// TIA Portal V20 export
Screen "Pop-up_Hmi_Opmodes18_h_Popup"  585x540
  ScreenItem "Background" at 0,0 size 585x540  Type=HmiRectangle
  ScreenItem "Dummy8" at 293,111 size 25x25  Type=HmiRectangle
  ScreenItem "Dummy9" at 319,111 size 25x25  Type=HmiRectangle
  ScreenItem "Dummy10" at 345,111 size 25x25  Type=HmiRectangle
  ScreenItem "Dummy11" at 371,111 size 25x25  Type=HmiRectangle
  ScreenItem "Dummy12" at 397,111 size 25x25  Type=HmiRectangle
  ScreenItem "Textfeld_1" at 77,106 size 29x30  Type=HmiTextBox
  ScreenItem "Dummy6" at 241,111 size 25x25  Type=HmiRectangle
  ScreenItem "Text_HmiPanelNo" at 244,50 size 160x23  Type=HmiTextBox
  ScreenItem "State_OPMode8_Select" at 293,80 size 25x25  Type=HmiTextBox
  ScreenItem "State_OPMode8_NotSelect" at 293,80 size 25x25  Type=HmiTextBox
  ScreenItem "State_OPMode8_Vis" at 293,80 size 25x25  Type=HmiRectangle
  ScreenItem "Descr_OPMode" at 108,26 size 305x20  Type=HmiTextBox
  ScreenItem "Dummy7" at 267,111 size 25x25  Type=HmiRectangle
  ScreenItem "Overview_OPMode" at 1,1 size 519x25  Type=HmiTextBox
  ScreenItem "State_OPMode1_Select" at 111,80 size 25x25  Type=HmiTextBox
  ScreenItem "State_OPMode1_NotSelect" at 111,80 size 25x25  Type=HmiTextBox
  ScreenItem "State_OPMode1_Vis" at 111,80 size 25x25  Type=HmiRectangle
  ScreenItem "State_OPMode2_Select" at 137,80 size 25x25  Type=HmiTextBox
  ScreenItem "State_OPMode2_NotSelect" at 137,80 size 25x25  Type=HmiTextBox
  ScreenItem "State_OPMode2_Vis" at 137,80 size 25x25  Type=HmiRectangle
  ScreenItem "State_OPMode3_Select" at 163,80 size 25x25  Type=HmiTextBox
  ScreenItem "State_OPMode3_NotSelect" at 163,80 size 25x25  Type=HmiTextBox
  ScreenItem "State_OPMode3_Vis" at 163,80 size 25x25  Type=HmiRectangle
  ScreenItem "State_OPMode4_Select" at 189,80 size 25x25  Type=HmiTextBox
  ScreenItem "State_OPMode4_NotSelect" at 189,80 size 25x25  Type=HmiTextBox
  ScreenItem "State_OPMode4_Vis" at 189,80 size 25x25  Type=HmiRectangle
  ScreenItem "State_OPMode5_Select" at 215,80 size 25x25  Type=HmiTextBox
  ScreenItem "State_OPMode5_NotSelect" at 215,80 size 25x25  Type=HmiTextBox
  ScreenItem "State_OPMode5_Vis" at 215,80 size 25x25  Type=HmiRectangle
  ScreenItem "State_OPMode6_Select" at 241,80 size 25x25  Type=HmiTextBox
  ScreenItem "State_OPMode6_NotSelect" at 241,80 size 25x25  Type=HmiTextBox
  ScreenItem "State_OPMode6_Vis" at 241,80 size 25x25  Type=HmiRectangle
  ScreenItem "State_OPMode7_Select" at 267,80 size 25x25  Type=HmiTextBox
  ScreenItem "State_OPMode7_NotSelect" at 267,80 size 25x25  Type=HmiTextBox
  ScreenItem "State_OPMode7_Vis" at 267,80 size 25x25  Type=HmiRectangle
  ScreenItem "State_OPMode9_Select" at 319,80 size 25x25  Type=HmiTextBox
  ScreenItem "State_OPMode9_NotSelect" at 319,80 size 25x25  Type=HmiTextBox
  ScreenItem "State_OPMode9_Vis" at 319,80 size 25x25  Type=HmiRectangle
  ScreenItem "State_OPMode10_Select" at 345,80 size 25x25  Type=HmiTextBox
  ScreenItem "State_OPMode10_NotSelect" at 345,80 size 25x25  Type=HmiTextBox
  ScreenItem "State_OPMode10_Vis" at 345,80 size 25x25  Type=HmiRectangle
  ScreenItem "State_OPMode11_Select" at 371,80 size 25x25  Type=HmiTextBox
  ScreenItem "State_OPMode11_NotSelect" at 371,80 size 25x25  Type=HmiTextBox
  ScreenItem "State_OPMode11_Vis" at 371,80 size 25x25  Type=HmiRectangle
  ScreenItem "State_OPMode12_Select" at 397,80 size 25x25  Type=HmiTextBox
  ScreenItem "State_OPMode12_NotSelect" at 397,80 size 25x25  Type=HmiTextBox
  ScreenItem "State_OPMode12_Vis" at 397,80 size 25x25  Type=HmiRectangle
  ScreenItem "Dummy13" at 424,111 size 25x25  Type=HmiRectangle
  ScreenItem "Dummy14" at 450,111 size 25x25  Type=HmiRectangle
  ScreenItem "Dummy15" at 476,111 size 25x25  Type=HmiRectangle
  ScreenItem "Dummy16" at 502,111 size 25x25  Type=HmiRectangle
  ScreenItem "Dummy17" at 528,111 size 25x25  Type=HmiRectangle
  ScreenItem "State_OPMode13_Select" at 424,80 size 25x25  Type=HmiTextBox
  ScreenItem "State_OPMode13_NotSelect" at 424,80 size 25x25  Type=HmiTextBox
  ScreenItem "State_OPMode13_Vis" at 424,80 size 25x25  Type=HmiRectangle
  ScreenItem "State_OPMode14_Select" at 450,80 size 25x25  Type=HmiTextBox
  ScreenItem "State_OPMode14_NotSelect" at 450,80 size 25x25  Type=HmiTextBox
  ScreenItem "State_OPMode14_Vis" at 450,80 size 25x25  Type=HmiRectangle
  ScreenItem "State_OPMode15_Select" at 476,80 size 25x25  Type=HmiTextBox
  ScreenItem "State_OPMode15_NotSelect" at 476,80 size 25x25  Type=HmiTextBox
  ScreenItem "State_OPMode15_Vis" at 476,80 size 25x25  Type=HmiRectangle
  ScreenItem "State_OPMode16_Select" at 502,80 size 25x25  Type=HmiTextBox
  ScreenItem "State_OPMode16_NotSelect" at 502,80 size 25x25  Type=HmiTextBox
  ScreenItem "State_OPMode16_Vis" at 502,80 size 25x25  Type=HmiRectangle
  ScreenItem "State_OPMode17_Select" at 528,80 size 25x25  Type=HmiTextBox
  ScreenItem "State_OPMode17_NotSelect" at 528,80 size 25x25  Type=HmiTextBox
  ScreenItem "State_OPMode17_Vis" at 528,80 size 25x25  Type=HmiRectangle
  ScreenItem "Dummy18" at 554,111 size 25x25  Type=HmiRectangle
  ScreenItem "State_OPMode18_Select" at 554,80 size 25x25  Type=HmiTextBox
  ScreenItem "State_OPMode18_NotSelect" at 554,80 size 25x25  Type=HmiTextBox
  ScreenItem "State_OPMode18_Vis" at 554,80 size 25x25  Type=HmiRectangle
  ScreenItem "Button_Back" at 1,1 size 90x60  Type=HmiButton
  ScreenItem "Button_Close" at 492,1 size 90x60  Type=HmiButton
  ScreenItem "Text_OPModeArea" at -84,288 size 260x25  Type=HmiTextBox
